(* IEC 61131-3 sources: axsharp/src/AXSharp.templates/working/templates/axsharpconsole/ax/src, 2 files *)

(* ---- configuration.st ---- *)
CONFIGURATION MyConfiguration
    TASK Main(Interval := T#10ms, Priority := 1);
    PROGRAM P1 WITH Main: MyProgram;

    VAR_GLOBAL
        Counter : ULINT;
    END_VAR
END_CONFIGURATION

(* ---- program.st ---- *)
PROGRAM MyProgram
    VAR_EXTERNAL
        Counter : ULINT;
    END_VAR

    Counter := Counter + ULINT#1;
END_PROGRAM
